(* IEC 61131-3 sources: trust-platform/crates/trust-runtime/tests/fixtures/oscat/oop_core/src, 1 file *)

(* ---- main.st ---- *)
PROGRAM Main
END_PROGRAM
